Universal Robots URScript: T002_qwen2.5-coder_32b_baseline_rep1_retry1.urscript

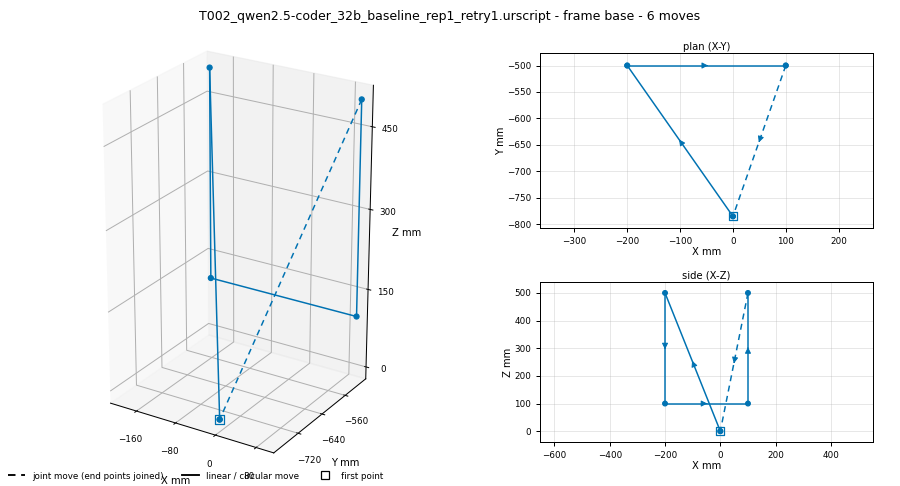
[picture p0: tool path of T002_qwen2.5-coder_32b_baseline_rep1_retry1.urscript in frame base, 6 of 6 moves have a stored position in this frame; points joined in program order, loops and branches not executed]
def linear_weld_path():
    # Go to home position
    movej(p[0.0, -0.785398, 0.0, -2.356194, 0.0, 0.0], a=1.2, v=1.0)

    # Approach above weld start
    movel(p[-0.2, -0.5, 0.5, -2.356194, 0.0, 0.0], a=1.2, v=0.25)

    # Descend to weld start position
    movel(p[-0.2, -0.5, 0.1, -2.356194, 0.0, 0.0], a=1.2, v=0.1)

    # Weld seam — 300mm linear path
    set_do(7,True)  # Activate welding arc
    movel(p[0.1, -0.5, 0.1, -2.356194, 0.0, 0.0], a=1.2, v=0.05)
    set_do(7,False)  # Deactivate welding arc

    # Retract above weld end
    movel(p[0.1, -0.5, 0.5, -2.356194, 0.0, 0.0], a=1.2, v=0.2)

    # Return to home position
    movej(p[0.0, -0.785398, 0.0, -2.356194, 0.0, 0.0], a=1.2, v=1.0)
end

# Execute the weld path function
linear_weld_path()
